(* IEC 61131-3 sources: trust-platform/examples/statechart_backend/src, 2 files *)

(* ---- config.st ---- *)
CONFIGURATION Config
RESOURCE MainResource ON PLC
    TASK MainTask (INTERVAL := T#10ms, PRIORITY := 1);
    PROGRAM P1 WITH MainTask : Main;
END_RESOURCE
VAR_CONFIG
    P1.DO0 AT %QX0.0 : BOOL;
    P1.DO1 AT %QX0.1 : BOOL;
    P1.DO2 AT %QX0.2 : BOOL;
    P1.DO3 AT %QX0.3 : BOOL;
    P1.DO4 AT %QX0.4 : BOOL;
    P1.DO5 AT %QX0.5 : BOOL;
    P1.DO6 AT %QX0.6 : BOOL;
    P1.DO7 AT %QX0.7 : BOOL;
END_VAR
END_CONFIGURATION

(* ---- Main.st ---- *)
(*
    Minimal ST program for StateChart hardware execution

    This program defines the I/O variables that will be controlled
    via the StateChart editor through the control endpoint.
*)

PROGRAM Main
VAR
    // Digital outputs mapped to EtherCAT EL2008
    DO0 : BOOL;
    DO1 : BOOL;
    DO2 : BOOL;
    DO3 : BOOL;
    DO4 : BOOL;
    DO5 : BOOL;
    DO6 : BOOL;
    DO7 : BOOL;

    // Heartbeat to show program is running
    heartbeat : BOOL;
END_VAR

// Toggle heartbeat every cycle
heartbeat := NOT heartbeat;

// Outputs are controlled via StateChart action mappings
// through the control endpoint, not by this program

END_PROGRAM
